Fanuc KAREL source: kb00097.KL

-- PROVISIONAL review KL for V1013-1; original PC SHA256 fe1a92bbc1fa71957f09a30a133a7044e5842f8597f9d7606d44eb81f35e2ca4
-- Incomplete behavior may be omitted. Consult companion uncertainty JSON. Do not deploy.
PROGRAM KB00097
%NOLOCKGROUP
BEGIN
  -- UNRESOLVED_PC offsets 5-14; opcodes 3F,75
  -- UNRESOLVED_PC offsets 19-26; opcodes 9D,23
  -- UNRESOLVED_PC offsets 31-38; opcodes 9D,23
  -- UNRESOLVED_PC offsets 43-50; opcodes 9D,23
  -- UNRESOLVED_PC offsets 55-64; opcodes 3F,75
  -- UNRESOLVED_PC offsets 69-76; opcodes 9D,23
  -- UNRESOLVED_PC offsets 81-125; opcodes 27,22,2A,22,22,22,22,2A,22,31
  -- UNRESOLVED_PC offsets 130-134; opcodes 7F
END KB00097
